(* IEC 61131-3 sources: llm-plc-st-eval/data/definitivo/qwen2.5-coder_14b/B5/zero_shot, 3 files *)

(* ---- ejec_1.st ---- *)
```pascal
FUNCTION_BLOCK FB_Ventilador
VAR_INPUT
    quemadorOn : BOOL; // Indica si el quemador está encendido
END_VAR

VAR_OUTPUT
    ventilador : BOOL; // Controla el ventilador
END_VAR

VAR
    timer : TON; // Timer de retardo
    timerDone : BOOL; // Indica si el timer ha terminado
END_VAR

// Inicialización del timer
IF NOT timerDone THEN
    timer(IN := NOT quemadorOn, PT := T#30S);
    timerDone := timer.Q;
END_IF;

// Control del ventilador
IF quemadorOn OR NOT timerDone THEN
    ventilador := TRUE;
ELSE
    ventilador := FALSE;
END_IF;
```

Este código implementa un FUNCTION_BLOCK llamado `FB_Ventilador` que controla el funcionamiento de un ventilador de enfriamiento en un horno. El ventilador se enciende cuando el quemador está encendido y continúa funcionando durante 30 segundos después de que el quemador se apague.

(* ---- ejec_2.st ---- *)
```pascal
FUNCTION_BLOCK FB_Ventilador
VAR_INPUT
    quemadorOn : BOOL; // Estado del quemador (TRUE si encendido, FALSE si apagado)
END_VAR

VAR_OUTPUT
    ventilador : BOOL; // Estado del ventilador (TRUE si encendido, FALSE si apagado)
END_VAR

VAR
    timer : TON; // Timer de retardo
    timerDone : BOOL; // Bandera para indicar si el timer ha terminado
END_VAR

// Inicialización del timer
IF NOT timerDone THEN
    timer(IN := NOT quemadorOn, PT := T#30S);
    timerDone := timer.Q;
END_IF;

// Control del ventilador
IF quemadorOn OR (NOT quemadorOn AND NOT timerDone) THEN
    ventilador := TRUE;
ELSE
    ventilador := FALSE;
END_IF;
```

Este código implementa un FUNCTION_BLOCK llamado `FB_Ventilador` que controla el funcionamiento de un ventilador de enfriamiento en un horno. El ventilador se enciende cuando el quemador está encendido y continúa funcionando durante 30 segundos después de que el quemador se apague.

(* ---- ejec_3.st ---- *)
```iec
FUNCTION_BLOCK FB_Ventilador
VAR_INPUT
    quemadorOn : BOOL; // Estado del quemador (encendido/apagado)
END_VAR

VAR_OUTPUT
    ventilador : BOOL; // Estado del ventilador (encendido/apagado)
END_VAR

VAR
    timer : TON; // Timer de retardo
    timerDone : BOOL; // Bandera para indicar que el timer ha terminado
END_VAR

// Inicialización del timer
IF NOT timer.Q THEN
    timer(IN := FALSE, PT := T#30S);
END_IF;

// Lógica del ventilador
IF quemadorOn THEN
    ventilador := TRUE; // El ventilador se enciende cuando el quemador está encendido
    timer(IN := FALSE); // Reinicia el timer
ELSE
    IF NOT timer.Q THEN
        timer(IN := TRUE); // Inicia el timer cuando el quemador se apaga
    END_IF;
    ventilador := timer.Q; // El ventilador se apaga cuando el timer termina
END_IF;
```

Este código implementa el comportamiento del ventilador de enfriamiento de un horno según las especificaciones proporcionadas. El ventilador se enciende cuando el quemador está encendido y continúa funcionando durante 30 segundos después de que el quemador se apaga.
